Fanuc KAREL source: kd00065.KL

-- PROVISIONAL review KL for V770-1; original PC SHA256 73423e4a65b8badb6988d78d5cca0f7c08f425b05730033cdb77b7e735c1cdef
-- Incomplete behavior may be omitted. Consult companion uncertainty JSON. Do not deploy.
PROGRAM KD00065
%NOLOCKGROUP
VAR
  I : INTEGER
  J : INTEGER
  B : BOOLEAN
  R : REAL
  S : STRING[80]
BEGIN
  -- UNRESOLVED_PC offsets 5-17; opcodes 9D,81,18,9D,1B,9D,12,13,04
  -- UNRESOLVED_PC offsets 22-26; opcodes 7F
END KD00065
